Staubli VAL3: utRectangle.pjx

--- utRectangle.pjx ---
Parameters version=s8.10.2Cs9_BS1991 stackSize=5000 millimeterUnit=true
Program file=start.pgx
Program file=stop.pgx
Data file=utRectangle.dtx
Type name=utBorder path=./utBorder/utBorder.pjx
Type name=utAppearance path=./utAppearance/utAppearance.pjx
Type name=utCommon path=./utCommon/utCommon.pjx
Type name=utText path=./utText/utText.pjx

--- utRectangle.dtx ---
public utBorder Border
  [0]
    string sBorderColour
    string sBorderWidth
public utAppearance Appearance
  [0]
    string sBackgroundColour
    string sColour
    bool bVisibility
public utCommon Common
  [0]
    bool bDisabled
    string sValue
    string sID
    num nValue
    string sPage
public utText Text
  [0]
    string sFontFamily
    string sFontStyle
    string sFontWeight
    string sTextAlignment
    num nFontSize

--- start.pgx ---
program start()
begin
end

--- stop.pgx ---
program stop()
begin
end
